// TIA Portal V19 export
TYPE "AnaMon.Status"
   STRUCT
      PV : Real;
      PV_unit : Int;
      PV_HiAlm : Bool;
      PV_HiWrn : Bool;
      PV_LoWrn : Bool;
      PV_LoAlm : Bool;
      MsgSup : Bool;
   END_STRUCT;
END_TYPE
